FUNCTION_BLOCK BasicAdapter (* Adapter communication, events only *)
  (* Standard: 61499-1 Annex A; Description: Copyright (c) 2023 Johannes Kepler University Linz This program and the accompanying materials are made available under the terms of the Eclipse Public License 2.0 which is available at https://www.eclipse.org/legal/epl-2.0/ SPDX-License-Identifier: EPL-2.0 *)
  (* Version 1.0, 2023-03-08, Bianca Wiesmayr, Johannes Kepler University Linz, initial API and implementation and/or initial documentation *)
  (* Documentation:
  ch
  *)
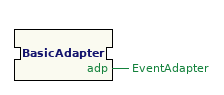
  PLUGS
    adp : EventAdapter;
  END_PLUGS
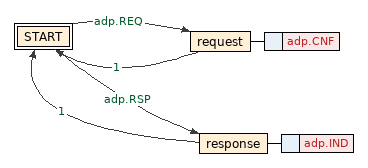
  EC_STATES
    START; (* Initial State *)
    request : -> adp.CNF;
    response : -> adp.IND;
  END_STATES
  EC_TRANSITIONS
    START TO request := adp.REQ;
    request TO START := 1;
    START TO response := adp.RSP;
    response TO START := 1;
  END_TRANSITIONS
END_FUNCTION_BLOCK
